Universal Robots URScript: MAIN_1.script

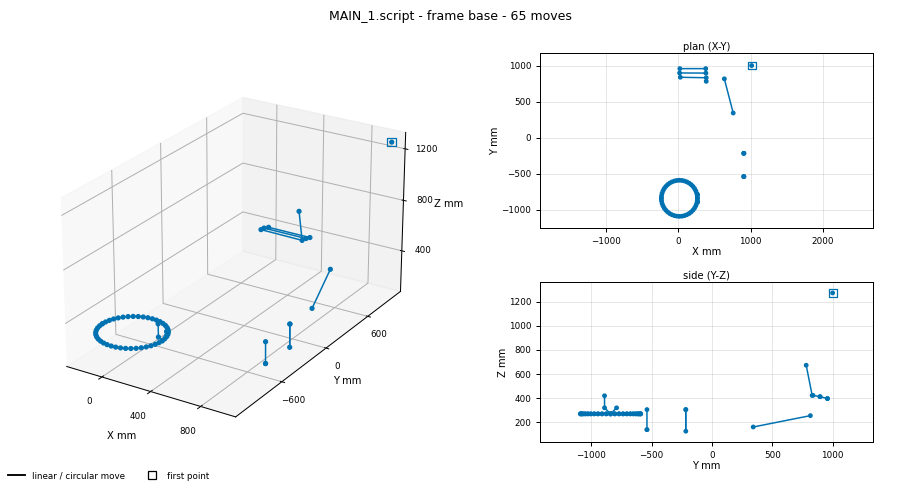
[picture p0: tool path of MAIN_1.script in frame base, 65 of 76 moves have a stored position in this frame; points joined in program order, loops and branches not executed]
def MAIN_1():
  # Global parameters:
  global speed_ms    = 0.250
  global speed_rads  = 0.750
  global accel_mss   = 1.200
  global accel_radss = 1.200
  global blend_radius_m = 0.001
  global ref_frame = p[0,0,0,0,0,0]

  #
  # TO REMOVE HEADER:
  # Go to "Program" -> "Post-Processor Editor"
  # Select "Universal Robots"
  # Set "INCLUDE_HEADER" to "False"
  #
  #--------------------------
  # Add any default subprograms here
  # For example, to drive a gripper as a program call:
  # def Gripper_Open():
  #   ...
  # end
  #
  # Example to drive a spray gun:
  def SprayOn(value):
    # use the value as an output:
    DO_SPRAY = 5
    if value == 0:
      set_standard_digital_out(DO_SPRAY, False)
    else:
      set_standard_digital_out(DO_SPRAY, True)
    end
  end

  # Example to drive an extruder:
  def Extruder(value):
    # use the value as an output:
    if value < 0:
      # stop extruder
    else:
      # start extruder
    end
  end

  # Example to move an external axis
  def MoveAxis(value):
    # use the value as an output:
    DO_AXIS_1 = 1
    DI_AXIS_1 = 1
    if value <= 0:
      set_standard_digital_out(DO_AXIS_1, False)

      # Wait for digital input to change state
      #while (get_standard_digital_in(DI_AXIS_1) != False):
      #  sync()
      #end
    else:
      set_standard_digital_out(DO_AXIS_1, True)

      # Wait for digital input to change state
      #while (get_standard_digital_in(DI_AXIS_1) != True):
      #  sync()
      #end
    end
  end
  #--------------------------

  # Subprogram PROG1_withaverylongnameandspecialcharacters
  def PROG1_withaverylongnameandspecialcharacters():
    # This is a subprogram call to PROG_1
    ref_frame = p[0.000000, 1.000000, 0.000000, 0.000000, 0.000000, 0.000000]
    set_tcp(p[0.000000, 0.000000, 0.200000, 0.000000, 0.000000, 0.000000])
    movej([-0.000000, 0.000000, 0.000000, 0.000000, 0.000000, -0.000000],accel_radss,speed_rads,0,0.001)
  end


  # Main program:
  # Program generated by RoboDK v5.6.9 for RoboDK Industrial on 26/02/2024 09:58:20
  # Using nominal kinematics.
  movej([-0.000000, 0.000000, 0.000000, 0.000000, 0.000000, -0.000000],accel_radss,speed_rads,0,0)
  movej([0.000000, 0.056047, -0.269194, 0.000000, 0.213148, -0.000000],accel_radss,speed_rads,0,0.001)
  movel(pose_trans(ref_frame,p[1.015000, 0.000000, 1.272000, 0.000000, 1.570796, 0.000000]),accel_mss,speed_ms,0,0) # end trace
  set_standard_digital_out(5, True)
  set_standard_digital_out(5, True)
  set_standard_digital_out(5, False)
  set_standard_digital_out(5, true)
  set_standard_analog_out(5, 1)
  set_standard_analog_out(5, 2)
  set_standard_analog_out(5, 0.5)
  set_standard_analog_out(5, true)
  var = val
  var = val
  while (get_standard_digital_in(5) != True):
    sync()
  end
  while (get_standard_digital_in(5) != True):
    sync()
  end
  while (get_standard_digital_in(5) != 0.5):
    sync()
  end
  while (get_standard_digital_in(5) != true):
    sync()
  end
  while (get_standard_digital_in(5) != True):
    sync()
  end
  while (var != val):
    sync()
  end
  while (var != val):
    sync()
  end
  popup("Message","Message",False,False,blocking=False)
  REMOTE_PROG_CALL_171()
  CODE_INSERT_172
  # Insert Comment
  ref_frame = p[0.719013, -0.664003, 0.000000, 0.000000, 0.000000, 0.000000]
  set_tcp(p[0.129073, 0.000000, 0.085477, 0.000000, 0.398790, 0.000000])
  accel_radss = 13.963
  speed_rads  = 3.142
  blend_radius_m = 0.010
  movej([-0.511943, 0.814667, -0.000428, 0.463308, 0.443239, -0.901183],accel_radss,speed_rads,0,0.010)
  blend_radius_m = 0.000
  accel_mss   = 0.200
  speed_ms    = 0.100
  movel(pose_trans(ref_frame,p[0.187786, 0.125499, 0.139112, -0.000082, 3.138451, 0.000110]),accel_mss,speed_ms,0,0.000)
  set_standard_digital_out(5, True)
  PICK_PART_111()
  blend_radius_m = 0.010
  accel_mss   = 0.600
  speed_ms    = 0.300
  movel([-0.511943, 0.814667, -0.000427, 0.463312, 0.443239, -0.901187],accel_mss,speed_ms,0,0)
  movel(pose_trans(ref_frame,p[0.187272, 0.447522, 0.305347, 0.000027, 3.138364, -0.000055]),accel_mss,speed_ms,0,0.010)
  blend_radius_m = 0.000
  accel_mss   = 0.200
  speed_ms    = 0.100
  # MoveSearch command not implemented
  movel(pose_trans(ref_frame,p[0.187851, 0.447517, 0.126235, 0.000027, 3.138364, -0.000055]),accel_mss,speed_ms,0,0.000)
  set_standard_digital_out(5, False)
  PLACE_PART_112()
  blend_radius_m = 0.010
  movel(pose_trans(ref_frame,p[0.187272, 0.447522, 0.305347, 0.000027, 3.138364, -0.000055]),accel_mss,speed_ms,0,0.010)
  ref_frame = p[0.577670, 0.392250, 0.000000, 0.000000, 0.000000, 0.679972]
  blend_radius_m = 0.025
  accel_radss = 13.963
  speed_rads  = 3.142
  accel_mss   = 0.200
  movej([0.910818, 0.797193, 0.120777, 1.164732, 0.347884, -1.618444],accel_radss,speed_rads,0,0.025)
  movec(pose_trans(ref_frame,p[0.430047, 0.043774, 0.231503, -1.148259, 2.734445, 0.138099]),pose_trans(ref_frame,p[0.109688, -0.153222, 0.161073, -1.148259, 2.734445, 0.138099]),accel_mss,speed_ms,0.025)
  # Circular movement using joint targets is not supported. Change the target type to cartesian or use a joint movement.
  blend_radius_m = 0.000
  accel_mss   = 0.200
  movel(pose_trans(ref_frame,p[0.312208, 0.292214, 0.255156, -1.148259, 2.734445, 0.138099]),accel_mss,speed_ms,0,0.000)
  movej([-0.000000, 0.000000, 0.000000, 0.000000, 0.000000, -0.000000],accel_radss,speed_rads,0,0)
  ref_frame = p[0.000000, 0.782714, 0.377610, 0.000000, 0.000000, 0.000000]
  movej([1.547688, 0.516645, -0.112204, -0.034631, 0.863575, 0.079372],accel_radss,speed_rads,0,0.000)
  movel(pose_trans(ref_frame,p[0.019898, 0.174307, 0.019008, 2.079600, -2.265750, 0.107759]),accel_mss,speed_ms,0,0.000)
  movel(pose_trans(ref_frame,p[0.378402, 0.174416, 0.018997, 2.079600, -2.265750, 0.107759]),accel_mss,speed_ms,0,0.000)
  movel(pose_trans(ref_frame,p[0.380996, 0.112363, 0.034882, 1.963520, -2.143933, 0.343573]),accel_mss,speed_ms,0,0.000)
  movel(pose_trans(ref_frame,p[0.016551, 0.114359, 0.034226, 1.963520, -2.143933, 0.343573]),accel_mss,speed_ms,0,0.000)
  movel(pose_trans(ref_frame,p[0.026434, 0.054524, 0.046072, -2.078092, 2.285598, 0.087159]),accel_mss,speed_ms,0,0.000)
  movel(pose_trans(ref_frame,p[0.385448, 0.048050, 0.045137, -2.018705, 2.221797, 0.218488]),accel_mss,speed_ms,0,0.000)
  movel(pose_trans(ref_frame,p[0.385448, -0.001625, 0.295251, -2.018705, 2.221797, 0.218488]),accel_mss,speed_ms,0,0.000)
  movej([-0.000000, 0.000000, 0.000000, 0.000000, 0.000000, -0.000000],accel_radss,speed_rads,0,0)
  EVENT_PROG_START_101()
  blend_radius_m = 0.001
  speed_ms    = 1.000
  ref_frame = p[0.013637, -0.840080, 0.000000, 0.000000, 0.000000, -1.570796]
  # Show Tool 1
  movej([-1.188400, 0.422403, 0.467495, 0.666950, 0.631839, -1.724322],accel_radss,speed_rads,0,0) # end trace
  EVENT_PATH_APPROACH_102()
  movel(pose_trans(ref_frame,p[-0.049895, 0.253259, 0.319999, -2.218137, 2.218140, 0.006349]),accel_mss,speed_ms,0,0.001)
  movel(pose_trans(ref_frame,p[0.000000, 0.250000, 0.270000, -2.218137, 2.218140, 0.006349]),accel_mss,speed_ms,0,0) # end trace
  EVENT_PATH_START_103()
  speed_ms    = 0.050
  movel(pose_trans(ref_frame,p[0.035579, 0.247455, 0.270000, -2.217769, 2.217778, 0.005226]),accel_mss,speed_ms,0,0.001)
  movel(pose_trans(ref_frame,p[0.070433, 0.239873, 0.270000, -2.217481, 2.217457, 0.004006]),accel_mss,speed_ms,0,0.001)
  movel(pose_trans(ref_frame,p[0.103854, 0.227408, 0.270000, -2.217271, 2.217250, 0.002728]),accel_mss,speed_ms,0,0.001)
  movel(pose_trans(ref_frame,p[0.135160, 0.210313, 0.270000, -2.217131, 2.217112, 0.001374]),accel_mss,speed_ms,0,0.001)
  movel(pose_trans(ref_frame,p[0.163715, 0.188937, 0.270000, -2.217087, 2.217069, 0.000000]),accel_mss,speed_ms,0,0.001)
  movel(pose_trans(ref_frame,p[0.188937, 0.163715, 0.270000, -2.217131, 2.217112, -0.001374]),accel_mss,speed_ms,0,0.001)
  movel(pose_trans(ref_frame,p[0.210313, 0.135160, 0.270000, -2.217254, 2.217233, -0.002728]),accel_mss,speed_ms,0,0.001)
  movel(pose_trans(ref_frame,p[0.227408, 0.103854, 0.270000, -2.217473, 2.217448, -0.004025]),accel_mss,speed_ms,0,0.001)
  movel(pose_trans(ref_frame,p[0.239873, 0.070433, 0.270000, -2.217760, 2.217769, -0.005245]),accel_mss,speed_ms,0,0.001)
  movel(pose_trans(ref_frame,p[0.247455, 0.035579, 0.270000, -2.218137, 2.218140, -0.006349]),accel_mss,speed_ms,0,0.001)
  movel(pose_trans(ref_frame,p[0.250000, 0.000000, 0.270000, -2.218575, 2.218572, -0.007318]),accel_mss,speed_ms,0,0.001)
  movel(pose_trans(ref_frame,p[0.247455, -0.035579, 0.270000, -2.219073, 2.219065, -0.008153]),accel_mss,speed_ms,0,0.001)
  movel(pose_trans(ref_frame,p[0.239873, -0.070433, 0.270000, -2.219605, 2.219630, -0.008833]),accel_mss,speed_ms,0,0.001)
  movel(pose_trans(ref_frame,p[0.227408, -0.103854, 0.270000, -2.220191, 2.220212, -0.009319]),accel_mss,speed_ms,0,0.001)
  movel(pose_trans(ref_frame,p[0.210313, -0.135160, 0.270000, -2.220802, 2.220821, -0.009593]),accel_mss,speed_ms,0,0.001)
  movel(pose_trans(ref_frame,p[0.188937, -0.163715, 0.270000, -2.221422, 2.221440, -0.009693]),accel_mss,speed_ms,0,0.001)
  movel(pose_trans(ref_frame,p[0.163715, -0.188937, 0.270000, 2.220802, -2.220821, 0.009593]),accel_mss,speed_ms,0,0.001)
  movel(pose_trans(ref_frame,p[0.135160, -0.210313, 0.270000, 2.220191, -2.220212, 0.009319]),accel_mss,speed_ms,0,0.001)
  movel(pose_trans(ref_frame,p[0.103854, -0.227408, 0.270000, 2.219605, -2.219630, 0.008833]),accel_mss,speed_ms,0,0.001)
  movel(pose_trans(ref_frame,p[0.070433, -0.239873, 0.270000, 2.219073, -2.219065, 0.008153]),accel_mss,speed_ms,0,0.001)
  movel(pose_trans(ref_frame,p[0.035579, -0.247455, 0.270000, 2.218575, -2.218572, 0.007318]),accel_mss,speed_ms,0,0.001)
  movel(pose_trans(ref_frame,p[0.000000, -0.250000, 0.270000, 2.218575, -2.218572, 0.007318]),accel_mss,speed_ms,0,0.001)
  movel(pose_trans(ref_frame,p[0.000000, -0.250000, 0.270000, 2.218137, -2.218140, 0.006349]),accel_mss,speed_ms,0,0.001)
  movel(pose_trans(ref_frame,p[-0.035579, -0.247455, 0.270000, 2.217760, -2.217769, 0.005245]),accel_mss,speed_ms,0,0.001)
  movel(pose_trans(ref_frame,p[-0.070433, -0.239873, 0.270000, 2.217481, -2.217457, 0.004006]),accel_mss,speed_ms,0,0.001)
  movel(pose_trans(ref_frame,p[-0.103854, -0.227408, 0.270000, 2.217271, -2.217250, 0.002728]),accel_mss,speed_ms,0,0.001)
  movel(pose_trans(ref_frame,p[-0.135160, -0.210313, 0.270000, 2.217131, -2.217112, 0.001374]),accel_mss,speed_ms,0,0.001)
  movel(pose_trans(ref_frame,p[-0.163715, -0.188937, 0.270000, 2.217087, -2.217069, 0.000000]),accel_mss,speed_ms,0,0.001)
  movel(pose_trans(ref_frame,p[-0.188937, -0.163715, 0.270000, 2.217131, -2.217112, -0.001374]),accel_mss,speed_ms,0,0.001)
  movel(pose_trans(ref_frame,p[-0.210313, -0.135160, 0.270000, 2.217271, -2.217250, -0.002728]),accel_mss,speed_ms,0,0.001)
  movel(pose_trans(ref_frame,p[-0.227408, -0.103854, 0.270000, 2.217490, -2.217465, -0.004025]),accel_mss,speed_ms,0,0.001)
  movel(pose_trans(ref_frame,p[-0.239873, -0.070433, 0.270000, 2.217760, -2.217769, -0.005245]),accel_mss,speed_ms,0,0.001)
  movel(pose_trans(ref_frame,p[-0.247455, -0.035579, 0.270000, 2.218137, -2.218140, -0.006349]),accel_mss,speed_ms,0,0.001)
  movel(pose_trans(ref_frame,p[-0.250000, 0.000000, 0.270000, 2.218575, -2.218572, -0.007318]),accel_mss,speed_ms,0,0.001)
  movel(pose_trans(ref_frame,p[-0.247455, 0.035579, 0.270000, 2.219082, -2.219073, -0.008133]),accel_mss,speed_ms,0,0.001)
  movel(pose_trans(ref_frame,p[-0.239873, 0.070433, 0.270000, 2.219605, -2.219630, -0.008794]),accel_mss,speed_ms,0,0.001)
  movel(pose_trans(ref_frame,p[-0.227408, 0.103854, 0.270000, 2.220191, -2.220212, -0.009319]),accel_mss,speed_ms,0,0.001)
  movel(pose_trans(ref_frame,p[-0.210313, 0.135160, 0.270000, 2.220802, -2.220821, -0.009593]),accel_mss,speed_ms,0,0.001)
  movel(pose_trans(ref_frame,p[-0.188937, 0.163715, 0.270000, -2.221422, 2.221440, 0.009693]),accel_mss,speed_ms,0,0.001)
  movel(pose_trans(ref_frame,p[-0.163715, 0.188937, 0.270000, -2.220802, 2.220821, 0.009593]),accel_mss,speed_ms,0,0.001)
  movel(pose_trans(ref_frame,p[-0.135160, 0.210313, 0.270000, -2.220191, 2.220212, 0.009281]),accel_mss,speed_ms,0,0.001)
  movel(pose_trans(ref_frame,p[-0.103854, 0.227408, 0.270000, -2.219605, 2.219630, 0.008833]),accel_mss,speed_ms,0,0.001)
  movel(pose_trans(ref_frame,p[-0.070433, 0.239873, 0.270000, -2.219073, 2.219065, 0.008153]),accel_mss,speed_ms,0,0.001)
  movel(pose_trans(ref_frame,p[-0.035579, 0.247455, 0.270000, -2.218575, 2.218572, 0.007318]),accel_mss,speed_ms,0,0.001)
  movel(pose_trans(ref_frame,p[0.000000, 0.250000, 0.270000, -2.218575, 2.218572, 0.007318]),accel_mss,speed_ms,0,0) # end trace
  speed_ms    = 1.000
  EVENT_PATH_FINISH_105()
  movel(pose_trans(ref_frame,p[0.049895, 0.253258, 0.319999, -2.218575, 2.218572, 0.007318]),accel_mss,speed_ms,0,0.001)
  movel(pose_trans(ref_frame,p[0.049939, 0.252642, 0.419997, -2.218575, 2.218572, 0.007318]),accel_mss,speed_ms,0,0) # end trace
  EVENT_PATH_RETRACT_106()
  EVENT_PROG_FINISH_107()
  ref_frame = p[0.719013, -0.664003, 0.000000, 0.000000, 0.000000, 0.000000]
  movej([-0.511943, 0.814667, -0.000428, 0.463308, 0.443239, -0.901183],accel_radss,speed_rads,0,0.001)
  sleep(1.250)
  movel(pose_trans(ref_frame,p[0.187786, 0.125499, 0.139112, -0.000082, 3.138451, 0.000110]),accel_mss,speed_ms,0,0) # end trace
  while (get_standard_digital_in(1) != True):
    sync()
  end
  movel(pose_trans(ref_frame,p[0.187264, 0.125487, 0.305356, 0.000000, 3.138381, -0.000000]),accel_mss,speed_ms,0,0) # end trace
  PROG1_withaverylongnameandspecialcharacters()
  # End of main program
end

MAIN_1()
